// TIA Portal V20 export
// export: Created 2026-10-20T12:49:39.4296533Z, ExportSetting WithDefaults, DisplayName Totally Integrated Automation Portal, DisplayVersion V20 Update 6, DisplayName TIA Portal Openness, DisplayVersion V20 Update 6, DisplayName TIA Portal Version Control Interface, DisplayVersion V20 Update 6, DisplayName SINAMICS Startdrive Advanced, DisplayVersion V20 SP1, DisplayName SINAMICS Startdrive G130, G150, S120, S150, SINAMICS MV, G220, S200, S210, DisplayVersion V20 SP1, DisplayName SINAMICS Startdrive G110M, G120, G120C, G120D, G120P, G115D, DisplayVersion V20 SP1, DisplayName STEP 7 Professional, DisplayVersion V20 Update 6, DisplayName STEP 7 Safety, DisplayVersion V20 Update 2, DisplayName WinCC Basic/Comfort/Advanced, DisplayVersion V20 Update 6, DisplayName WinCC Unified, DisplayVersion V20 Update 6
DATA_BLOCK "Sf_C3204_FB_DB"   // DB276
VERSION : 0.1
// stored: AutoNumber true, DBAccessibleFromOPCUA true, InstanceOfName Safety_Stops_FB, InstanceOfType FB
"Safety_Stops_FB"
   // VAR_INPUT
   //    Sys_No : UInt;
   //    Mode : UInt;
   //    Timeout : UInt;
   //    Reset : Bool;
   // END_VAR
   // VAR_IN_OUT
   //    Sfts_Control : "Sfts_Control";
   // END_VAR
   // VAR
   //    State : UInt;
   //    LP_Timer { ExternalAccessible := 'False'; ExternalVisible := 'False'; ExternalWritable := 'False'} : TON_TIME;
   //    T_Run { S7_SetPoint := 'True'} : TOF_TIME;
   //    Timer_1 : Time;
   // END_VAR
BEGIN
END_DATA_BLOCK
